{attribute 'qualified_only'}
VAR_GLOBAL
	fbSFC_Temp1: FB_SFC_Template;
END_VAR

(* stored: Version 1.1.0.1, ProductVersion 3.1.4024.12
   GVL g_SFC: Id {60949f43-4a61-4329-b7c7-78e679279bde} *)
